Staubli VAL3: click_Stop.pgx

program click_Stop()
  local bool l_bResult
begin
  //立即停止机器人
  l_bResult=userPageConfirm("确认立即停止机器人？")
  if l_bResult
    rs:bToStopCycle=true
    delay(0.2)
    rs:bToStopCycle=false
  endIf
end
